(* IEC 61131-3 sources: SemantiST/compiler/toolchain/compatibility/profiles/codesys-conversions, 1 file *)

(* ---- conversions.st ---- *)
(* Generated by compiler/toolchain/compatibility/profiles/generate_codesys.py
   from the pinned RuSTy standard library. Do not edit by hand.
   CODESYS conversions the pinned RuSTy lacks, composed from RuSTy
   conversions with CODESYS semantics (low bits kept on narrowing, REAL
   rounded half away from zero, BOOL TRUE = 1). *)

FUNCTION BOOL_TO_REAL : REAL
VAR_INPUT IN : BOOL; END_VAR
    IF IN THEN
        BOOL_TO_REAL := 1.0;
    ELSE
        BOOL_TO_REAL := 0.0;
    END_IF;
END_FUNCTION

FUNCTION BOOL_TO_LREAL : LREAL
VAR_INPUT IN : BOOL; END_VAR
    IF IN THEN
        BOOL_TO_LREAL := 1.0;
    ELSE
        BOOL_TO_LREAL := 0.0;
    END_IF;
END_FUNCTION

FUNCTION BYTE_TO_REAL : REAL
VAR_INPUT IN : BYTE; END_VAR
    BYTE_TO_REAL := IN;
END_FUNCTION

FUNCTION BYTE_TO_LREAL : LREAL
VAR_INPUT IN : BYTE; END_VAR
    BYTE_TO_LREAL := IN;
END_FUNCTION

FUNCTION WORD_TO_REAL : REAL
VAR_INPUT IN : WORD; END_VAR
    WORD_TO_REAL := IN;
END_FUNCTION

FUNCTION WORD_TO_LREAL : LREAL
VAR_INPUT IN : WORD; END_VAR
    WORD_TO_LREAL := IN;
END_FUNCTION

FUNCTION DWORD_TO_LREAL : LREAL
VAR_INPUT IN : DWORD; END_VAR
    DWORD_TO_LREAL := IN;
END_FUNCTION

FUNCTION LWORD_TO_REAL : REAL
VAR_INPUT IN : LWORD; END_VAR
    LWORD_TO_REAL := IN;
END_FUNCTION

FUNCTION SINT_TO_BOOL : BOOL
VAR_INPUT IN : SINT; END_VAR
    SINT_TO_BOOL := IN <> 0;
END_FUNCTION

FUNCTION USINT_TO_BOOL : BOOL
VAR_INPUT IN : USINT; END_VAR
    USINT_TO_BOOL := IN <> 0;
END_FUNCTION

FUNCTION INT_TO_BOOL : BOOL
VAR_INPUT IN : INT; END_VAR
    INT_TO_BOOL := IN <> 0;
END_FUNCTION

FUNCTION UINT_TO_BOOL : BOOL
VAR_INPUT IN : UINT; END_VAR
    UINT_TO_BOOL := IN <> 0;
END_FUNCTION

FUNCTION UDINT_TO_BOOL : BOOL
VAR_INPUT IN : UDINT; END_VAR
    UDINT_TO_BOOL := IN <> 0;
END_FUNCTION

FUNCTION ULINT_TO_BOOL : BOOL
VAR_INPUT IN : ULINT; END_VAR
    ULINT_TO_BOOL := IN <> 0;
END_FUNCTION

FUNCTION REAL_TO_BOOL : BOOL
VAR_INPUT IN : REAL; END_VAR
    REAL_TO_BOOL := IN <> 0.0;
END_FUNCTION

FUNCTION REAL_TO_BYTE : BYTE
VAR_INPUT IN : REAL; END_VAR
VAR v : LINT; END_VAR
    v := REAL_TO_LINT(IN);
    REAL_TO_BYTE := LINT_TO_BYTE(v);
END_FUNCTION

FUNCTION REAL_TO_WORD : WORD
VAR_INPUT IN : REAL; END_VAR
VAR v : LINT; END_VAR
    v := REAL_TO_LINT(IN);
    REAL_TO_WORD := LINT_TO_WORD(v);
END_FUNCTION

FUNCTION REAL_TO_LWORD : LWORD
VAR_INPUT IN : REAL; END_VAR
VAR v : LINT; END_VAR
    v := REAL_TO_LINT(IN);
    REAL_TO_LWORD := LINT_TO_LWORD(v);
END_FUNCTION

FUNCTION LREAL_TO_BOOL : BOOL
VAR_INPUT IN : LREAL; END_VAR
    LREAL_TO_BOOL := IN <> 0.0;
END_FUNCTION

FUNCTION LREAL_TO_BYTE : BYTE
VAR_INPUT IN : LREAL; END_VAR
VAR v : LINT; END_VAR
    v := LREAL_TO_LINT(IN);
    LREAL_TO_BYTE := LINT_TO_BYTE(v);
END_FUNCTION

FUNCTION LREAL_TO_WORD : WORD
VAR_INPUT IN : LREAL; END_VAR
VAR v : LINT; END_VAR
    v := LREAL_TO_LINT(IN);
    LREAL_TO_WORD := LINT_TO_WORD(v);
END_FUNCTION

FUNCTION LREAL_TO_DWORD : DWORD
VAR_INPUT IN : LREAL; END_VAR
VAR v : LINT; END_VAR
    v := LREAL_TO_LINT(IN);
    LREAL_TO_DWORD := LINT_TO_DWORD(v);
END_FUNCTION

FUNCTION WORD_TO_STRING : STRING
VAR_INPUT IN : WORD; END_VAR
VAR v : ULINT; END_VAR
    v := IN;
    WORD_TO_STRING := ULINT_TO_STRING(v);
END_FUNCTION

FUNCTION SINT_TO_STRING : STRING
VAR_INPUT IN : SINT; END_VAR
VAR v : LINT; END_VAR
    v := IN;
    SINT_TO_STRING := LINT_TO_STRING(v);
END_FUNCTION

FUNCTION INT_TO_STRING : STRING
VAR_INPUT IN : INT; END_VAR
VAR v : LINT; END_VAR
    v := IN;
    INT_TO_STRING := LINT_TO_STRING(v);
END_FUNCTION

FUNCTION BOOL_TO_STRING : STRING
VAR_INPUT IN : BOOL; END_VAR
    IF IN THEN
        BOOL_TO_STRING := 'TRUE';
    ELSE
        BOOL_TO_STRING := 'FALSE';
    END_IF;
END_FUNCTION

FUNCTION STRING_TO_BYTE : BYTE
VAR_INPUT IN : STRING; END_VAR
    STRING_TO_BYTE := LINT_TO_BYTE(STRING_TO_LINT(IN));
END_FUNCTION

FUNCTION STRING_TO_WORD : WORD
VAR_INPUT IN : STRING; END_VAR
    STRING_TO_WORD := LINT_TO_WORD(STRING_TO_LINT(IN));
END_FUNCTION

FUNCTION STRING_TO_DWORD : DWORD
VAR_INPUT IN : STRING; END_VAR
    STRING_TO_DWORD := LINT_TO_DWORD(STRING_TO_LINT(IN));
END_FUNCTION

FUNCTION STRING_TO_LWORD : LWORD
VAR_INPUT IN : STRING; END_VAR
    STRING_TO_LWORD := LINT_TO_LWORD(STRING_TO_LINT(IN));
END_FUNCTION

FUNCTION STRING_TO_SINT : SINT
VAR_INPUT IN : STRING; END_VAR
    STRING_TO_SINT := LINT_TO_SINT(STRING_TO_LINT(IN));
END_FUNCTION

FUNCTION STRING_TO_USINT : USINT
VAR_INPUT IN : STRING; END_VAR
    STRING_TO_USINT := LINT_TO_USINT(STRING_TO_LINT(IN));
END_FUNCTION

FUNCTION STRING_TO_INT : INT
VAR_INPUT IN : STRING; END_VAR
    STRING_TO_INT := LINT_TO_INT(STRING_TO_LINT(IN));
END_FUNCTION

FUNCTION STRING_TO_UINT : UINT
VAR_INPUT IN : STRING; END_VAR
    STRING_TO_UINT := LINT_TO_UINT(STRING_TO_LINT(IN));
END_FUNCTION

FUNCTION STRING_TO_UDINT : UDINT
VAR_INPUT IN : STRING; END_VAR
    STRING_TO_UDINT := LINT_TO_UDINT(STRING_TO_LINT(IN));
END_FUNCTION

FUNCTION STRING_TO_ULINT : ULINT
VAR_INPUT IN : STRING; END_VAR
    STRING_TO_ULINT := LINT_TO_ULINT(STRING_TO_LINT(IN));
END_FUNCTION

FUNCTION __CDS_DWORD_TO_REAL : REAL
VAR_INPUT IN : DWORD; END_VAR
VAR v : ULINT; END_VAR
    v := IN;
    __CDS_DWORD_TO_REAL := ULINT_TO_REAL(v);
END_FUNCTION

FUNCTION __CDS_LREAL_TO_LWORD : LWORD
VAR_INPUT IN : LREAL; END_VAR
VAR v : LINT; END_VAR
    v := LREAL_TO_LINT(IN);
    __CDS_LREAL_TO_LWORD := LINT_TO_LWORD(v);
END_FUNCTION

FUNCTION __CDS_LWORD_TO_LREAL : LREAL
VAR_INPUT IN : LWORD; END_VAR
VAR v : ULINT; END_VAR
    v := IN;
    __CDS_LWORD_TO_LREAL := ULINT_TO_LREAL(v);
END_FUNCTION

FUNCTION __CDS_REAL_TO_DWORD : DWORD
VAR_INPUT IN : REAL; END_VAR
VAR v : LINT; END_VAR
    v := REAL_TO_LINT(IN);
    __CDS_REAL_TO_DWORD := LINT_TO_DWORD(v);
END_FUNCTION
